FUNCTION_BLOCK FB 500
VERSION : 0.1


VAR_INPUT
  IN0 : BOOL ;
  IN1 : BOOL ;
  IN2 : BOOL ;
END_VAR
VAR_OUTPUT
  OUT3 : BOOL ;
  OUT4 : BOOL ;
END_VAR
VAR
  STAT5 : BOOL ;
  STAT6 : BOOL ;
  STAT7 : BOOL ;
  STAT8 : BOOL ;
END_VAR
BEGIN
NETWORK
TITLE =
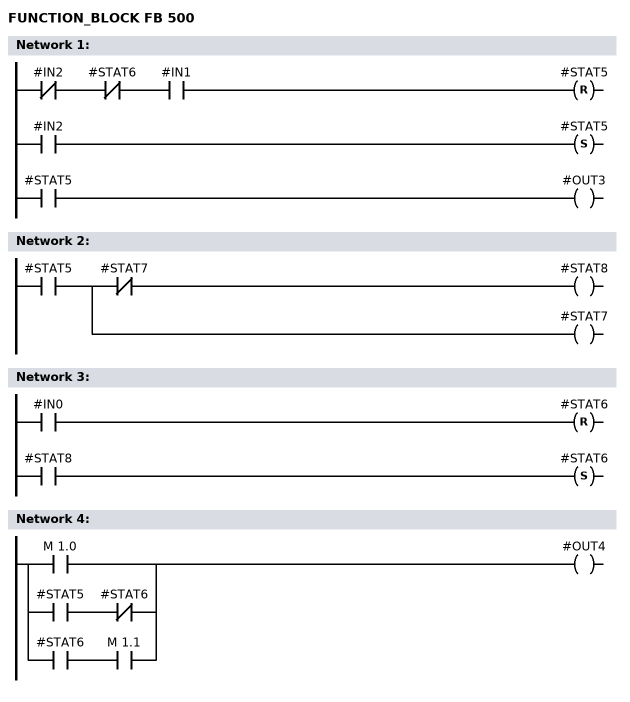

      AN    #IN2;
      AN    #STAT6;
      A     #IN1;
      R     #STAT5;
      A     #IN2;
      S     #STAT5;
      A     #STAT5;
      =     #OUT3;
NETWORK
TITLE =

      A     #STAT5;
      =     L      0.0;
      A     L      0.0;
      AN    #STAT7;
      =     #STAT8;
      A     L      0.0;
      BLD   102;
      =     #STAT7;
NETWORK
TITLE =

      A     #IN0;
      R     #STAT6;
      A     #STAT8;
      S     #STAT6;
      NOP   0;
NETWORK
TITLE =

      O     M      1.0;
      O     ;
      A     #STAT5;
      AN    #STAT6;
      O     ;
      A     #STAT6;
      A     M      1.1;
      =     #OUT4;
END_FUNCTION_BLOCK

FUNCTION FC 0 : VOID
VERSION : 0.1

BEGIN
NETWORK
TITLE =
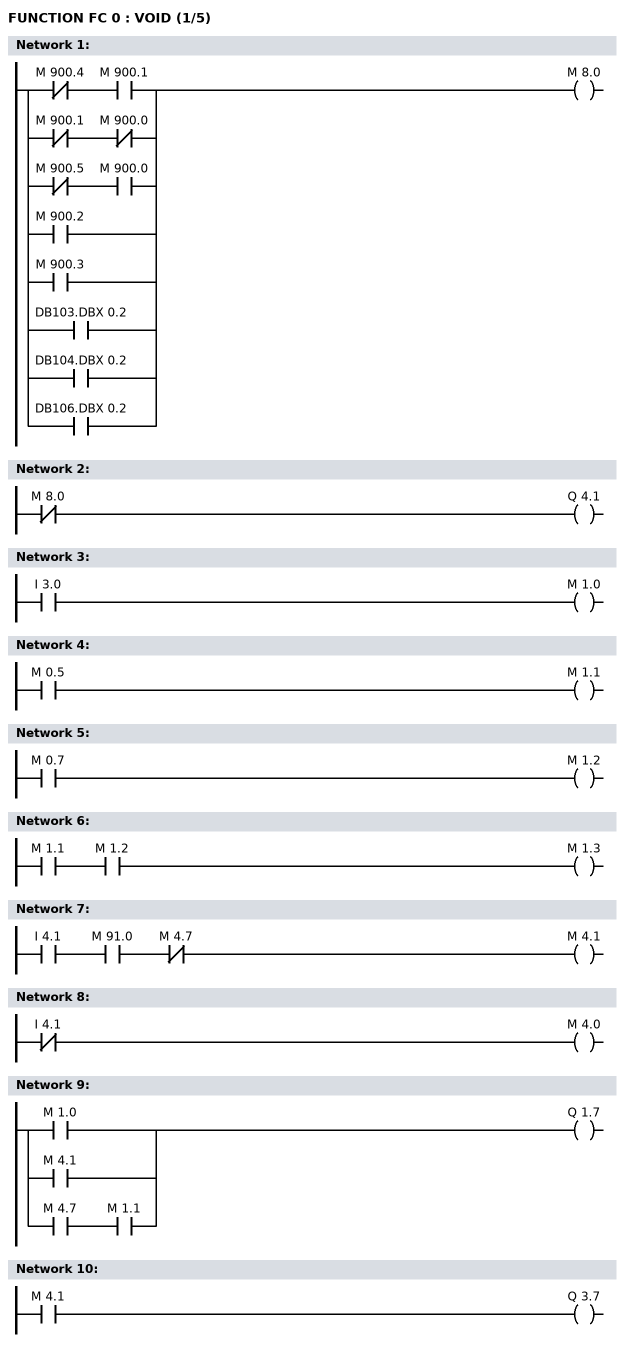

      AN    M    900.4;
      A     M    900.1;
      O     ;
      AN    M    900.1;
      AN    M    900.0;
      O     ;
      AN    M    900.5;
      A     M    900.0;
      O     M    900.2;
      O     M    900.3;
      O     DB103.DBX    0.2;
      O     DB104.DBX    0.2;
      O     DB106.DBX    0.2;
      =     M      8.0;
NETWORK
TITLE =

      AN    M      8.0;
      =     Q      4.1;
NETWORK
TITLE =

      A     I      3.0;
      =     M      1.0;
NETWORK
TITLE =

      A     M      0.5;
      =     M      1.1;
NETWORK
TITLE =

      A     M      0.7;
      =     M      1.2;
NETWORK
TITLE =

      A     M      1.1;
      A     M      1.2;
      =     M      1.3;
NETWORK
TITLE =

      A     I      4.1;
      A     M     91.0;
      AN    M      4.7;
      =     M      4.1;
NETWORK
TITLE =

      AN    I      4.1;
      =     M      4.0;
NETWORK
TITLE =

      O     M      1.0;
      O     M      4.1;
      O     ;
      A     M      4.7;
      A     M      1.1;
      =     Q      1.7;
NETWORK
TITLE =

      A     M      4.1;
      =     Q      3.7;
NETWORK
TITLE =
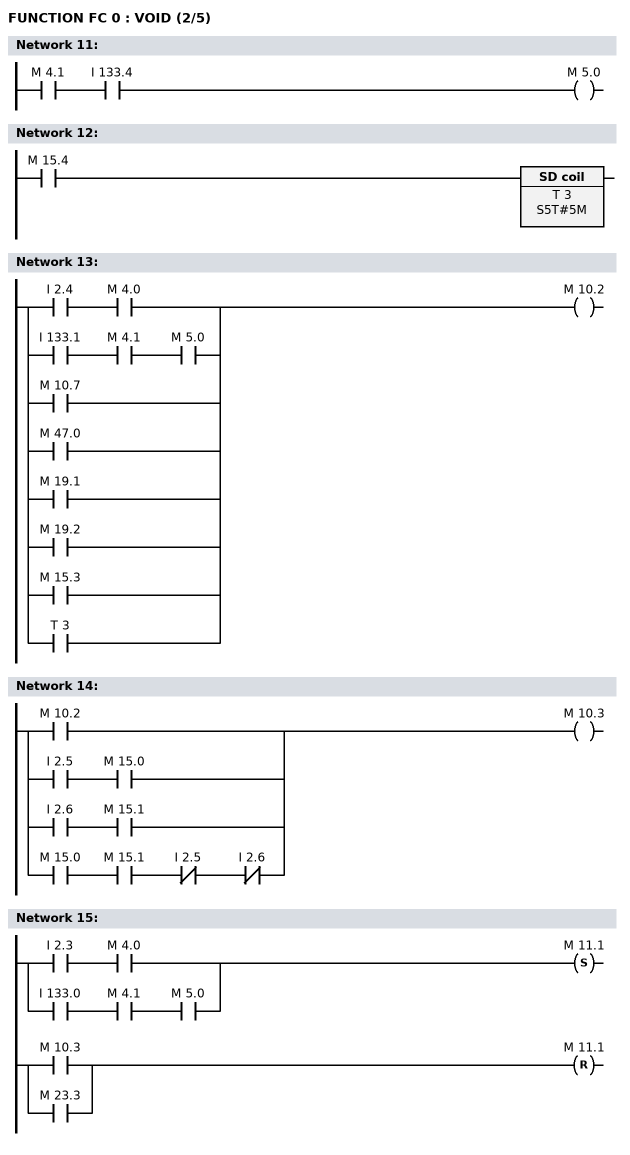

      A     M      4.1;
      A     I    133.4;
      =     M      5.0;
NETWORK
TITLE =

      A     M     15.4;
      L     S5T#5M;
      SD    T      3;
      NOP   0;
      NOP   0;
      NOP   0;
      NOP   0;
NETWORK
TITLE =

      A     I      2.4;
      A     M      4.0;
      O     ;
      A     I    133.1;
      A     M      4.1;
      A     M      5.0;
      O     M     10.7;
      O     M     47.0;
      O     M     19.1;
      O     M     19.2;
      O     M     15.3;
      O     T      3;
      =     M     10.2;
NETWORK
TITLE =

      O     M     10.2;
      O     ;
      A     I      2.5;
      A     M     15.0;
      O     ;
      A     I      2.6;
      A     M     15.1;
      O     ;
      A     M     15.0;
      A     M     15.1;
      AN    I      2.5;
      AN    I      2.6;
      =     M     10.3;
NETWORK
TITLE =

      A(    ;
      A     I      2.3;
      A     M      4.0;
      O     ;
      A     I    133.0;
      A     M      4.1;
      A     M      5.0;
      )     ;
      S     M     11.1;
      A(    ;
      O     M     10.3;
      O     M     23.3;
      )     ;
      R     M     11.1;
      NOP   0;
NETWORK
TITLE =
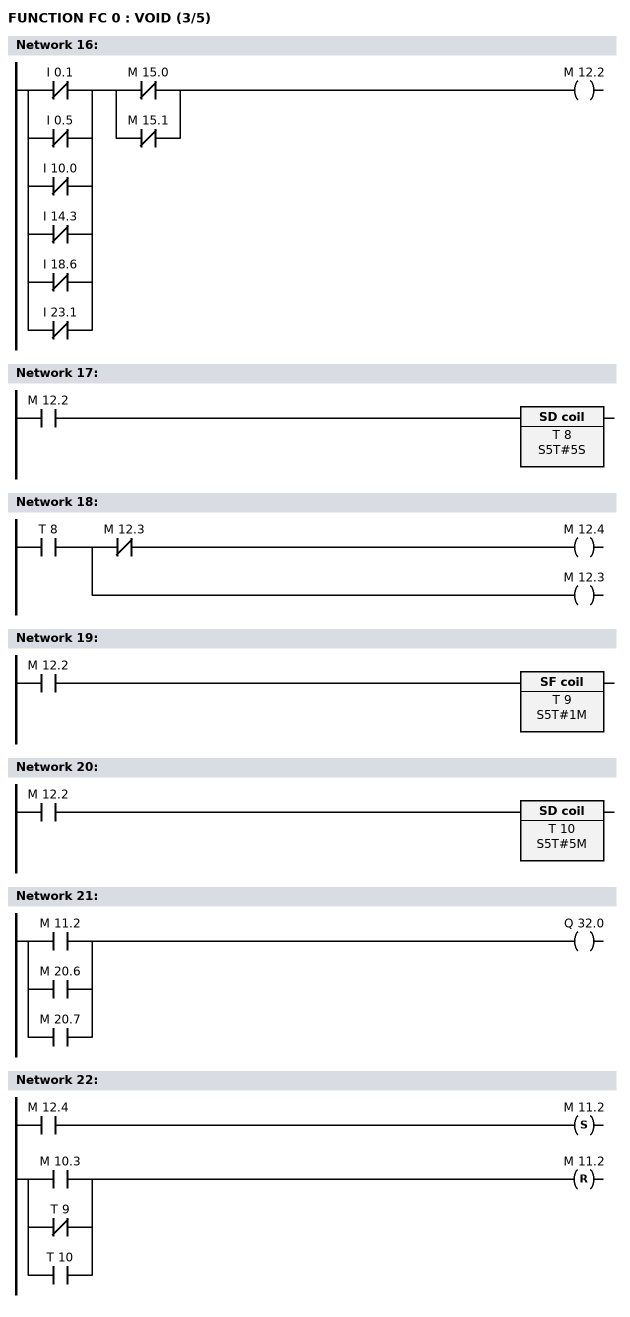

      A(    ;
      ON    I      0.1;
      ON    I      0.5;
      ON    I     10.0;
      ON    I     14.3;
      ON    I     18.6;
      ON    I     23.1;
      )     ;
      A(    ;
      ON    M     15.0;
      ON    M     15.1;
      )     ;
      =     M     12.2;
NETWORK
TITLE =

      A     M     12.2;
      L     S5T#5S;
      SD    T      8;
      NOP   0;
      NOP   0;
      NOP   0;
      NOP   0;
NETWORK
TITLE =

      A     T      8;
      =     L      0.0;
      A     L      0.0;
      AN    M     12.3;
      =     M     12.4;
      A     L      0.0;
      BLD   102;
      =     M     12.3;
NETWORK
TITLE =

      A     M     12.2;
      L     S5T#1M;
      SF    T      9;
      NOP   0;
      NOP   0;
      NOP   0;
      NOP   0;
NETWORK
TITLE =

      A     M     12.2;
      L     S5T#5M;
      SD    T     10;
      NOP   0;
      NOP   0;
      NOP   0;
      NOP   0;
NETWORK
TITLE =

      O     M     11.2;
      O     M     20.6;
      O     M     20.7;
      =     Q     32.0;
NETWORK
TITLE =

      A     M     12.4;
      S     M     11.2;
      A(    ;
      O     M     10.3;
      ON    T      9;
      O     T     10;
      )     ;
      R     M     11.2;
      NOP   0;
NETWORK
TITLE =
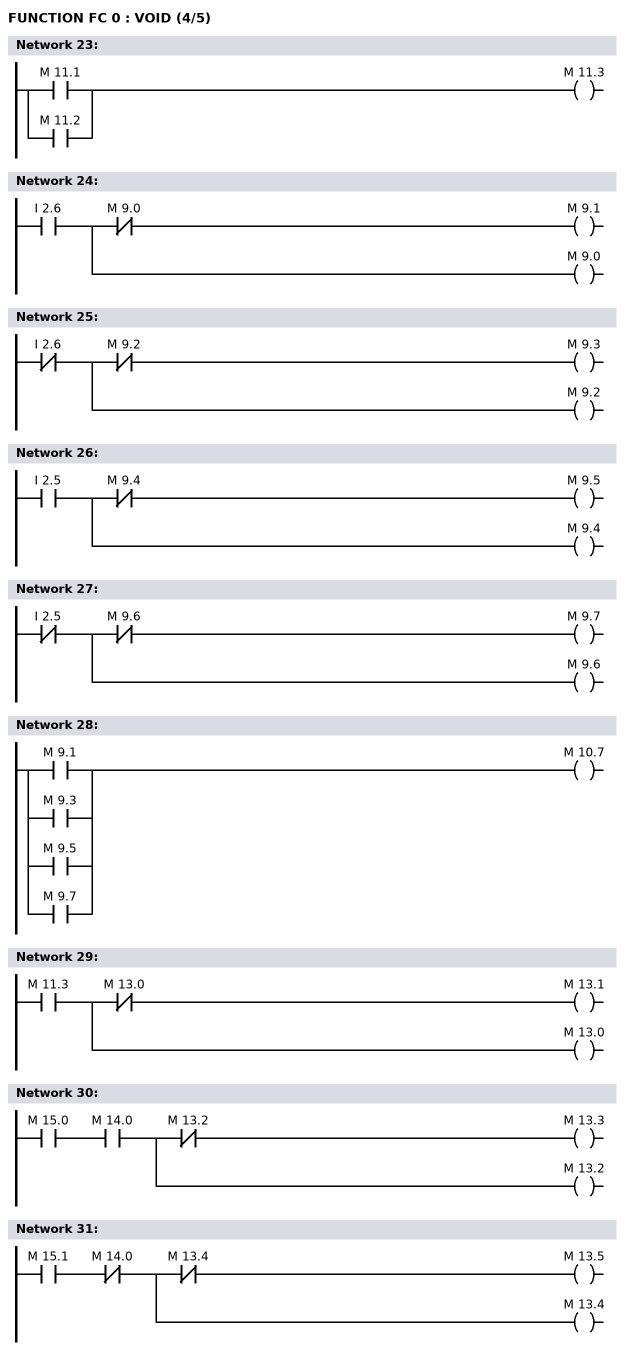

      O     M     11.1;
      O     M     11.2;
      =     M     11.3;
NETWORK
TITLE =

      A     I      2.6;
      =     L      0.0;
      A     L      0.0;
      AN    M      9.0;
      =     M      9.1;
      A     L      0.0;
      BLD   102;
      =     M      9.0;
NETWORK
TITLE =

      AN    I      2.6;
      =     L      0.0;
      A     L      0.0;
      AN    M      9.2;
      =     M      9.3;
      A     L      0.0;
      BLD   102;
      =     M      9.2;
NETWORK
TITLE =

      A     I      2.5;
      =     L      0.0;
      A     L      0.0;
      AN    M      9.4;
      =     M      9.5;
      A     L      0.0;
      BLD   102;
      =     M      9.4;
NETWORK
TITLE =

      AN    I      2.5;
      =     L      0.0;
      A     L      0.0;
      AN    M      9.6;
      =     M      9.7;
      A     L      0.0;
      BLD   102;
      =     M      9.6;
NETWORK
TITLE =

      O     M      9.1;
      O     M      9.3;
      O     M      9.5;
      O     M      9.7;
      =     M     10.7;
NETWORK
TITLE =

      A     M     11.3;
      =     L      0.0;
      A     L      0.0;
      AN    M     13.0;
      =     M     13.1;
      A     L      0.0;
      BLD   102;
      =     M     13.0;
NETWORK
TITLE =

      A     M     15.0;
      A     M     14.0;
      =     L      0.0;
      A     L      0.0;
      AN    M     13.2;
      =     M     13.3;
      A     L      0.0;
      BLD   102;
      =     M     13.2;
NETWORK
TITLE =

      A     M     15.1;
      AN    M     14.0;
      =     L      0.0;
      A     L      0.0;
      AN    M     13.4;
      =     M     13.5;
      A     L      0.0;
      BLD   102;
      =     M     13.4;
NETWORK
TITLE =
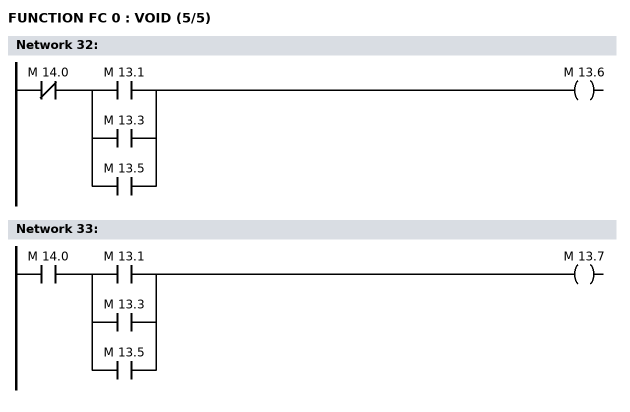

      AN    M     14.0;
      A(    ;
      O     M     13.1;
      O     M     13.3;
      O     M     13.5;
      )     ;
      =     M     13.6;
NETWORK
TITLE =

      A     M     14.0;
      A(    ;
      O     M     13.1;
      O     M     13.3;
      O     M     13.5;
      )     ;
      =     M     13.7;
NETWORK
TITLE =

      A(    ;
      A     M     13.7;
      R     M     14.0;
      A     M     13.6;
      S     M     14.0;
      A     M     14.0;
      )     ;
      AN    I      2.5;
      AN    I      2.6;
      O     I      2.5;
      =     M     14.2;
NETWORK
TITLE =
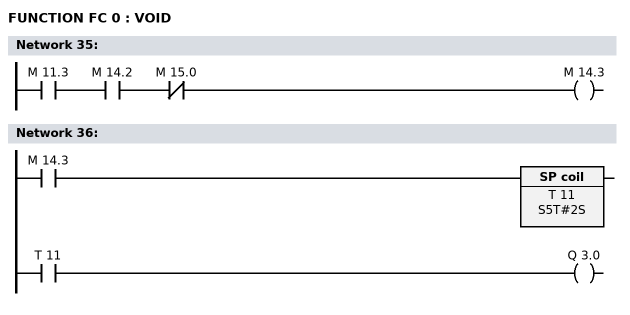

      A     M     11.3;
      A     M     14.2;
      AN    M     15.0;
      =     M     14.3;
NETWORK
TITLE =

      A     M     14.3;
      L     S5T#2S;
      SP    T     11;
      NOP   0;
      NOP   0;
      NOP   0;
      A     T     11;
      =     Q      3.0;
NETWORK
TITLE =

      A(    ;
      AN    M     14.3;
      L     S5T#2S;
      SP    T     12;
      NOP   0;
      NOP   0;
      NOP   0;
      A     T     12;
      )     ;
      NOT   ;
      =     Q      3.1;
NETWORK
TITLE =
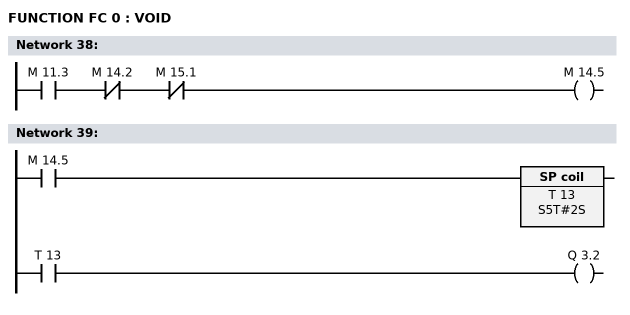

      A     M     11.3;
      AN    M     14.2;
      AN    M     15.1;
      =     M     14.5;
NETWORK
TITLE =

      A     M     14.5;
      L     S5T#2S;
      SP    T     13;
      NOP   0;
      NOP   0;
      NOP   0;
      A     T     13;
      =     Q      3.2;
NETWORK
TITLE =

      A(    ;
      AN    M     14.5;
      L     S5T#2S;
      SP    T     14;
      NOP   0;
      NOP   0;
      NOP   0;
      A     T     14;
      )     ;
      NOT   ;
      =     Q      3.3;
NETWORK
TITLE =
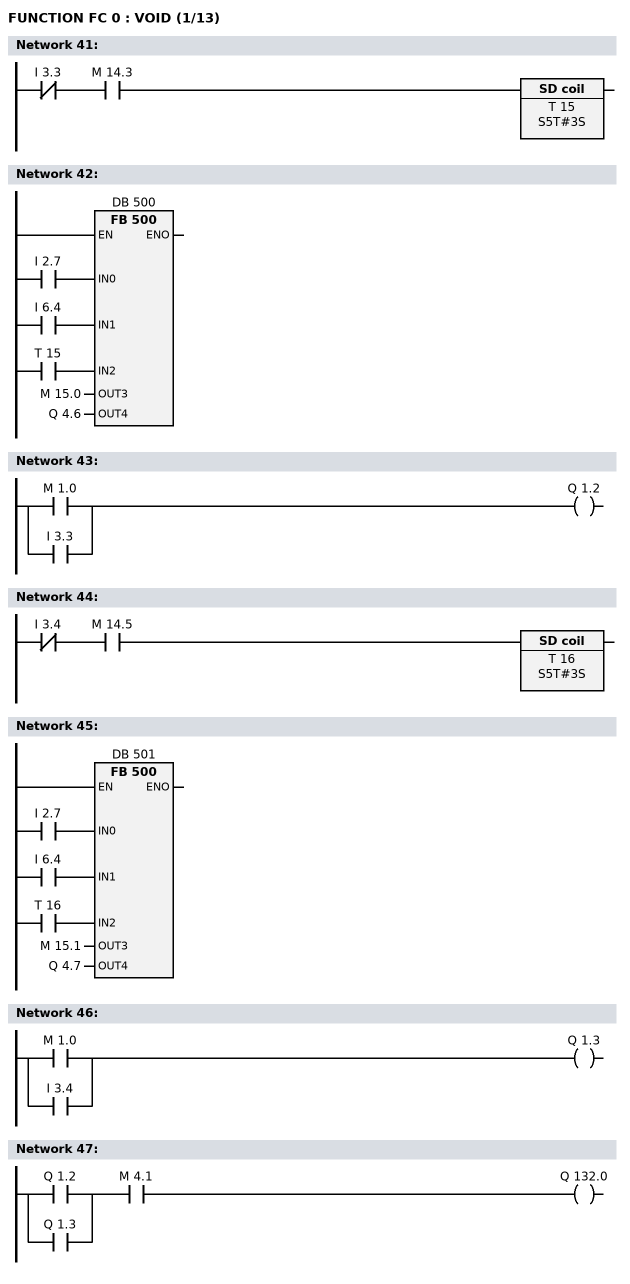

      AN    I      3.3;
      A     M     14.3;
      L     S5T#3S;
      SD    T     15;
      NOP   0;
      NOP   0;
      NOP   0;
      NOP   0;
NETWORK
TITLE =

      A     I      2.7;
      =     L      0.0;
      BLD   103;
      A     I      6.4;
      =     L      0.1;
      BLD   103;
      A     T     15;
      =     L      0.2;
      BLD   103;
      CALL FB   500 , DB   500 (
           IN0                      := L      0.0,
           IN1                      := L      0.1,
           IN2                      := L      0.2,
           OUT3                     := M     15.0,
           OUT4                     := Q      4.6);
      NOP   0;
NETWORK
TITLE =

      O     M      1.0;
      O     I      3.3;
      =     Q      1.2;
NETWORK
TITLE =

      AN    I      3.4;
      A     M     14.5;
      L     S5T#3S;
      SD    T     16;
      NOP   0;
      NOP   0;
      NOP   0;
      NOP   0;
NETWORK
TITLE =

      A     I      2.7;
      =     L      0.0;
      BLD   103;
      A     I      6.4;
      =     L      0.1;
      BLD   103;
      A     T     16;
      =     L      0.2;
      BLD   103;
      CALL FB   500 , DB   501 (
           IN0                      := L      0.0,
           IN1                      := L      0.1,
           IN2                      := L      0.2,
           OUT3                     := M     15.1,
           OUT4                     := Q      4.7);
      NOP   0;
NETWORK
TITLE =

      O     M      1.0;
      O     I      3.4;
      =     Q      1.3;
NETWORK
TITLE =

      A(    ;
      O     Q      1.2;
      O     Q      1.3;
      )     ;
      A     M      4.1;
      =     Q    132.0;
NETWORK
TITLE =
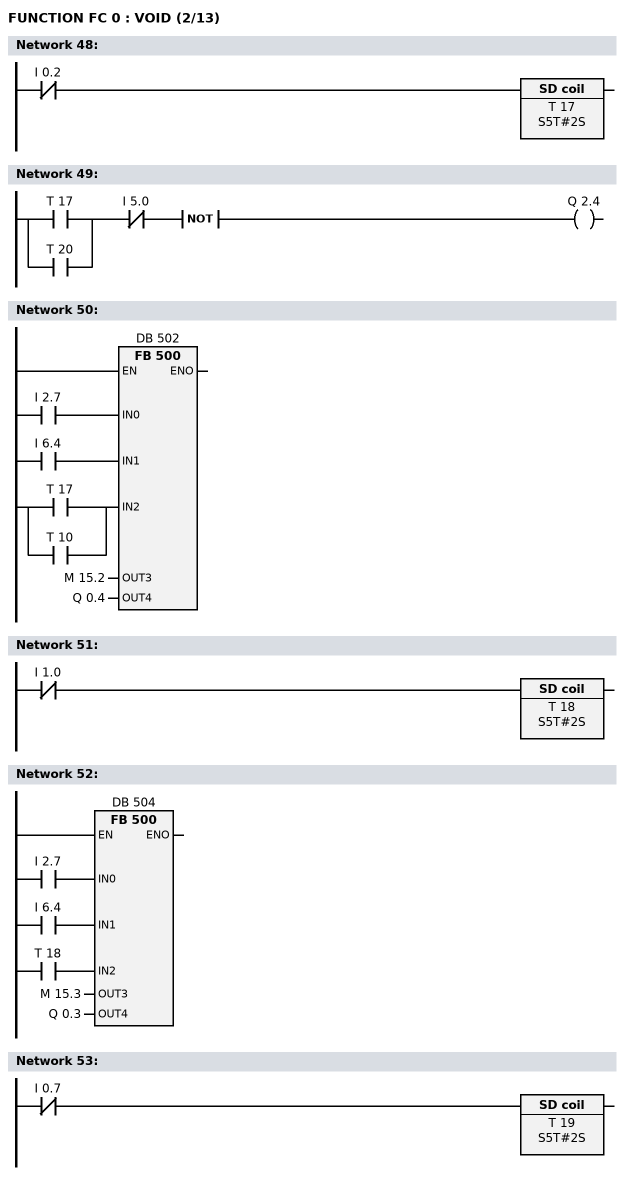

      AN    I      0.2;
      L     S5T#2S;
      SD    T     17;
      NOP   0;
      NOP   0;
      NOP   0;
      NOP   0;
NETWORK
TITLE =

      A(    ;
      O     T     17;
      O     T     20;
      )     ;
      AN    I      5.0;
      NOT   ;
      =     Q      2.4;
NETWORK
TITLE =

      A     I      2.7;
      =     L      0.0;
      BLD   103;
      A     I      6.4;
      =     L      0.1;
      BLD   103;
      A(    ;
      O     T     17;
      O     T     10;
      )     ;
      =     L      0.2;
      BLD   103;
      CALL FB   500 , DB   502 (
           IN0                      := L      0.0,
           IN1                      := L      0.1,
           IN2                      := L      0.2,
           OUT3                     := M     15.2,
           OUT4                     := Q      0.4);
      NOP   0;
NETWORK
TITLE =

      AN    I      1.0;
      L     S5T#2S;
      SD    T     18;
      NOP   0;
      NOP   0;
      NOP   0;
      NOP   0;
NETWORK
TITLE =

      A     I      2.7;
      =     L      0.0;
      BLD   103;
      A     I      6.4;
      =     L      0.1;
      BLD   103;
      A     T     18;
      =     L      0.2;
      BLD   103;
      CALL FB   500 , DB   504 (
           IN0                      := L      0.0,
           IN1                      := L      0.1,
           IN2                      := L      0.2,
           OUT3                     := M     15.3,
           OUT4                     := Q      0.3);
      NOP   0;
NETWORK
TITLE =

      AN    I      0.7;
      L     S5T#2S;
      SD    T     19;
      NOP   0;
      NOP   0;
      NOP   0;
      NOP   0;
NETWORK
TITLE =
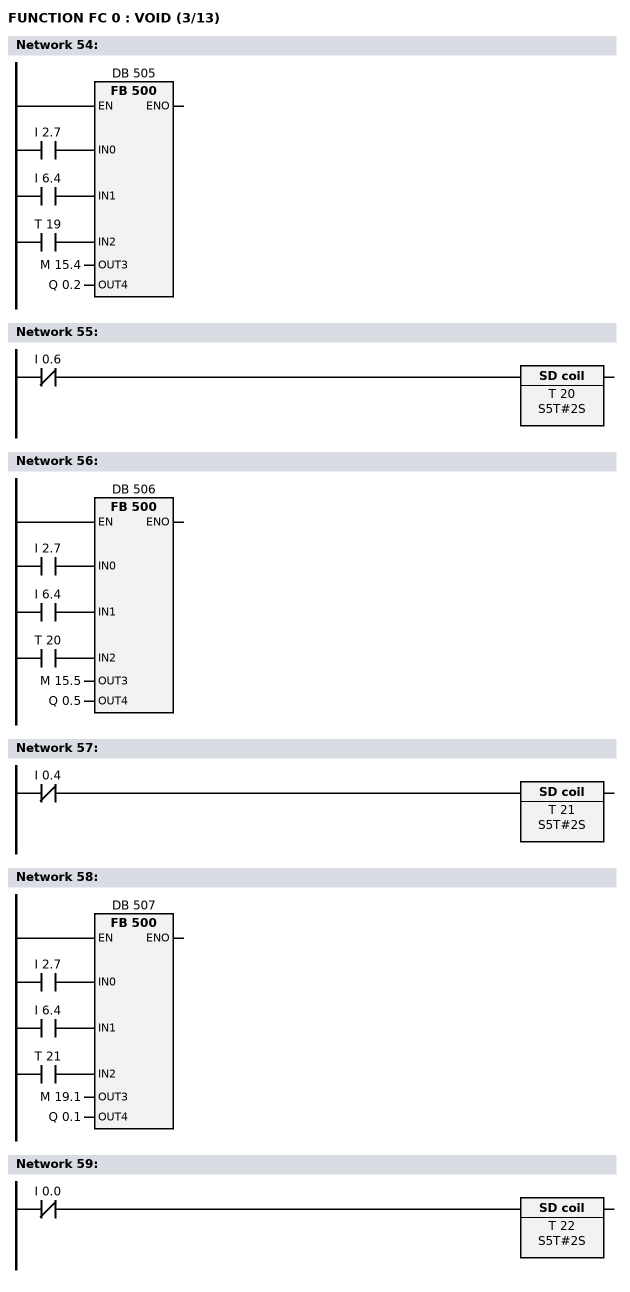

      A     I      2.7;
      =     L      0.0;
      BLD   103;
      A     I      6.4;
      =     L      0.1;
      BLD   103;
      A     T     19;
      =     L      0.2;
      BLD   103;
      CALL FB   500 , DB   505 (
           IN0                      := L      0.0,
           IN1                      := L      0.1,
           IN2                      := L      0.2,
           OUT3                     := M     15.4,
           OUT4                     := Q      0.2);
      NOP   0;
NETWORK
TITLE =

      AN    I      0.6;
      L     S5T#2S;
      SD    T     20;
      NOP   0;
      NOP   0;
      NOP   0;
      NOP   0;
NETWORK
TITLE =

      A     I      2.7;
      =     L      0.0;
      BLD   103;
      A     I      6.4;
      =     L      0.1;
      BLD   103;
      A     T     20;
      =     L      0.2;
      BLD   103;
      CALL FB   500 , DB   506 (
           IN0                      := L      0.0,
           IN1                      := L      0.1,
           IN2                      := L      0.2,
           OUT3                     := M     15.5,
           OUT4                     := Q      0.5);
      NOP   0;
NETWORK
TITLE =

      AN    I      0.4;
      L     S5T#2S;
      SD    T     21;
      NOP   0;
      NOP   0;
      NOP   0;
      NOP   0;
NETWORK
TITLE =

      A     I      2.7;
      =     L      0.0;
      BLD   103;
      A     I      6.4;
      =     L      0.1;
      BLD   103;
      A     T     21;
      =     L      0.2;
      BLD   103;
      CALL FB   500 , DB   507 (
           IN0                      := L      0.0,
           IN1                      := L      0.1,
           IN2                      := L      0.2,
           OUT3                     := M     19.1,
           OUT4                     := Q      0.1);
      NOP   0;
NETWORK
TITLE =

      AN    I      0.0;
      L     S5T#2S;
      SD    T     22;
      NOP   0;
      NOP   0;
      NOP   0;
      NOP   0;
NETWORK
TITLE =
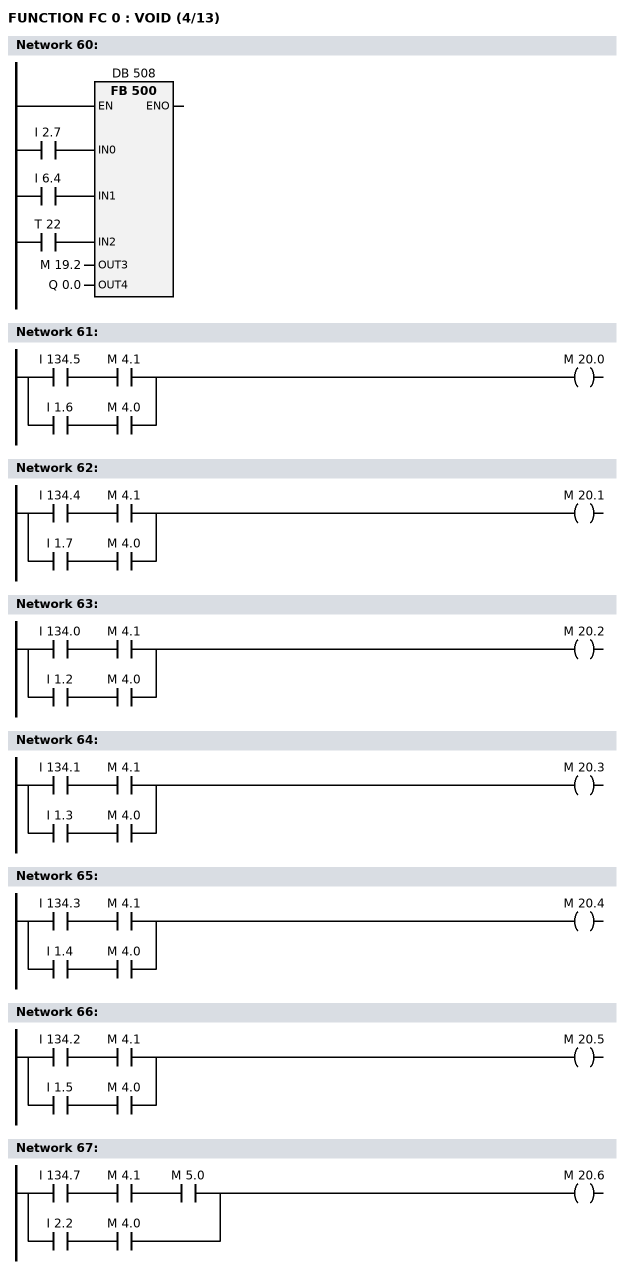

      A     I      2.7;
      =     L      0.0;
      BLD   103;
      A     I      6.4;
      =     L      0.1;
      BLD   103;
      A     T     22;
      =     L      0.2;
      BLD   103;
      CALL FB   500 , DB   508 (
           IN0                      := L      0.0,
           IN1                      := L      0.1,
           IN2                      := L      0.2,
           OUT3                     := M     19.2,
           OUT4                     := Q      0.0);
      NOP   0;
NETWORK
TITLE =

      A     I    134.5;
      A     M      4.1;
      O     ;
      A     I      1.6;
      A     M      4.0;
      =     M     20.0;
NETWORK
TITLE =

      A     I    134.4;
      A     M      4.1;
      O     ;
      A     I      1.7;
      A     M      4.0;
      =     M     20.1;
NETWORK
TITLE =

      A     I    134.0;
      A     M      4.1;
      O     ;
      A     I      1.2;
      A     M      4.0;
      =     M     20.2;
NETWORK
TITLE =

      A     I    134.1;
      A     M      4.1;
      O     ;
      A     I      1.3;
      A     M      4.0;
      =     M     20.3;
NETWORK
TITLE =

      A     I    134.3;
      A     M      4.1;
      O     ;
      A     I      1.4;
      A     M      4.0;
      =     M     20.4;
NETWORK
TITLE =

      A     I    134.2;
      A     M      4.1;
      O     ;
      A     I      1.5;
      A     M      4.0;
      =     M     20.5;
NETWORK
TITLE =

      A     I    134.7;
      A     M      4.1;
      A     M      5.0;
      O     ;
      A     I      2.2;
      A     M      4.0;
      =     M     20.6;
NETWORK
TITLE =
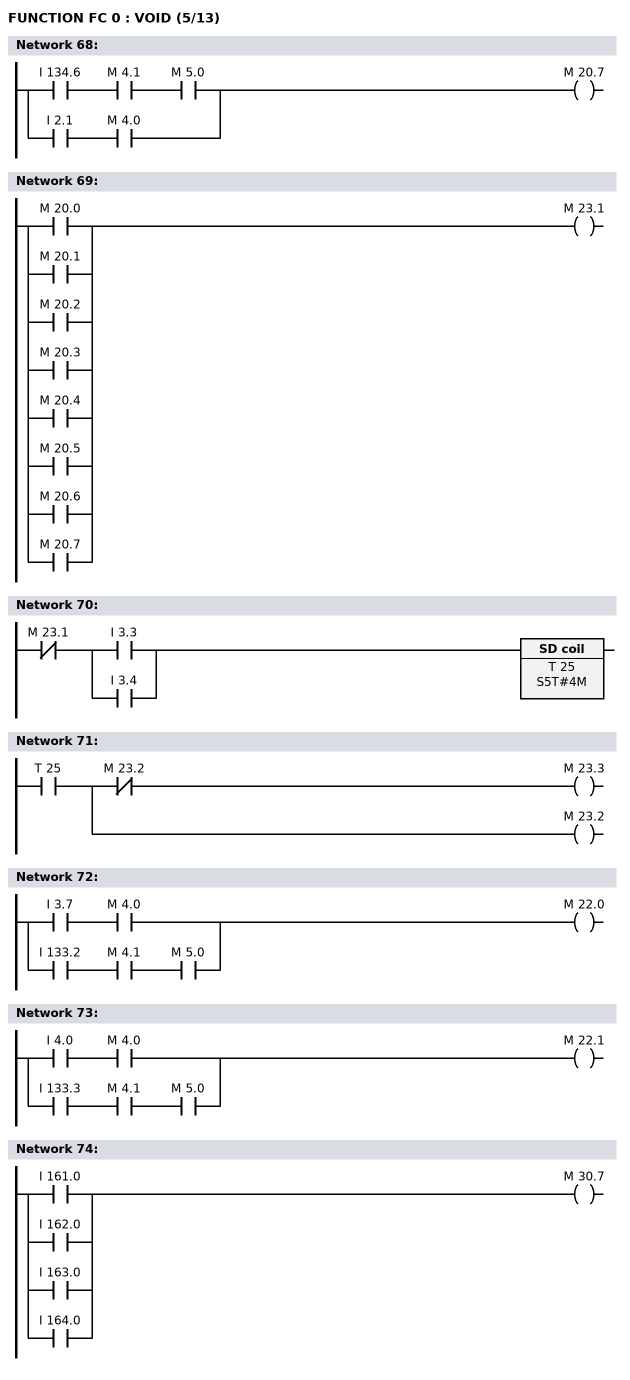

      A     I    134.6;
      A     M      4.1;
      A     M      5.0;
      O     ;
      A     I      2.1;
      A     M      4.0;
      =     M     20.7;
NETWORK
TITLE =

      O     M     20.0;
      O     M     20.1;
      O     M     20.2;
      O     M     20.3;
      O     M     20.4;
      O     M     20.5;
      O     M     20.6;
      O     M     20.7;
      =     M     23.1;
NETWORK
TITLE =

      AN    M     23.1;
      A(    ;
      O     I      3.3;
      O     I      3.4;
      )     ;
      L     S5T#4M;
      SD    T     25;
      NOP   0;
      NOP   0;
      NOP   0;
      NOP   0;
NETWORK
TITLE =

      A     T     25;
      =     L      0.0;
      A     L      0.0;
      AN    M     23.2;
      =     M     23.3;
      A     L      0.0;
      BLD   102;
      =     M     23.2;
NETWORK
TITLE =

      A     I      3.7;
      A     M      4.0;
      O     ;
      A     I    133.2;
      A     M      4.1;
      A     M      5.0;
      =     M     22.0;
NETWORK
TITLE =

      A     I      4.0;
      A     M      4.0;
      O     ;
      A     I    133.3;
      A     M      4.1;
      A     M      5.0;
      =     M     22.1;
NETWORK
TITLE =

      O     I    161.0;
      O     I    162.0;
      O     I    163.0;
      O     I    164.0;
      =     M     30.7;
NETWORK
TITLE =
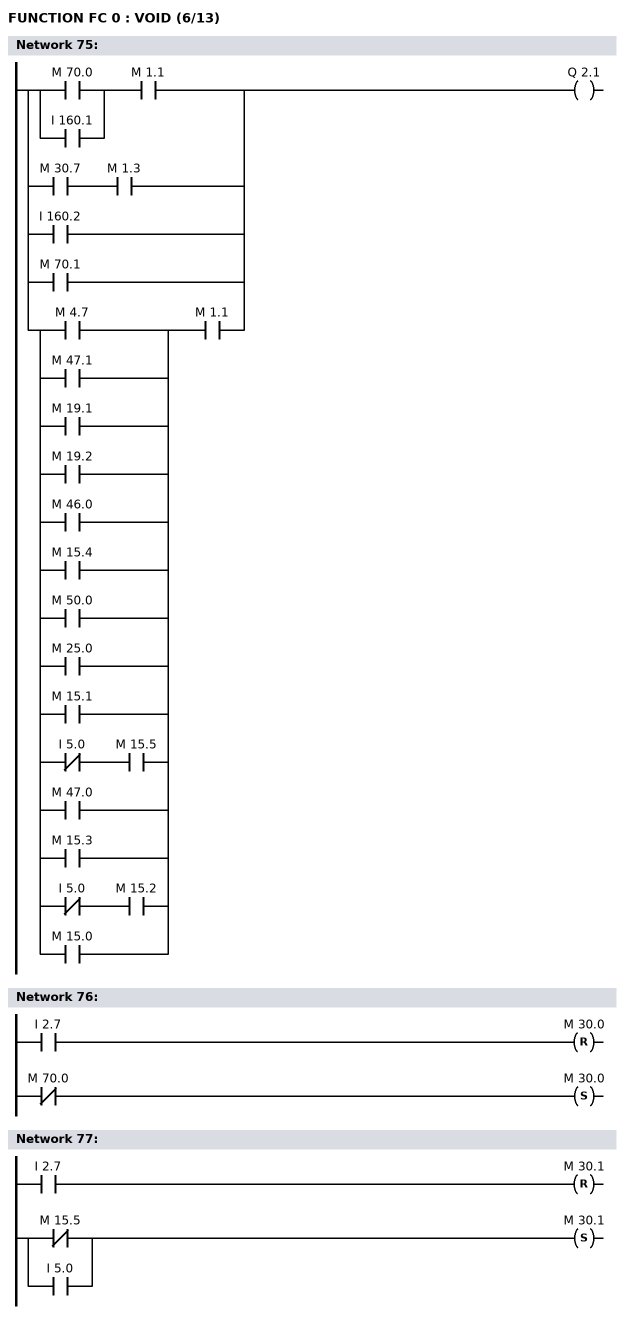

      A(    ;
      O     M     70.0;
      O     I    160.1;
      )     ;
      A     M      1.1;
      O     ;
      A     M     30.7;
      A     M      1.3;
      O     I    160.2;
      O     M     70.1;
      O     ;
      A(    ;
      O     M      4.7;
      O     M     47.1;
      O     M     19.1;
      O     M     19.2;
      O     M     46.0;
      O     M     15.4;
      O     M     50.0;
      O     M     25.0;
      O     M     15.1;
      O     ;
      AN    I      5.0;
      A     M     15.5;
      O     M     47.0;
      O     M     15.3;
      O     ;
      AN    I      5.0;
      A     M     15.2;
      O     M     15.0;
      )     ;
      A     M      1.1;
      =     Q      2.1;
NETWORK
TITLE =

      A     I      2.7;
      R     M     30.0;
      AN    M     70.0;
      S     M     30.0;
      NOP   0;
NETWORK
TITLE =

      A     I      2.7;
      R     M     30.1;
      A(    ;
      ON    M     15.5;
      O     I      5.0;
      )     ;
      S     M     30.1;
      NOP   0;
NETWORK
TITLE =
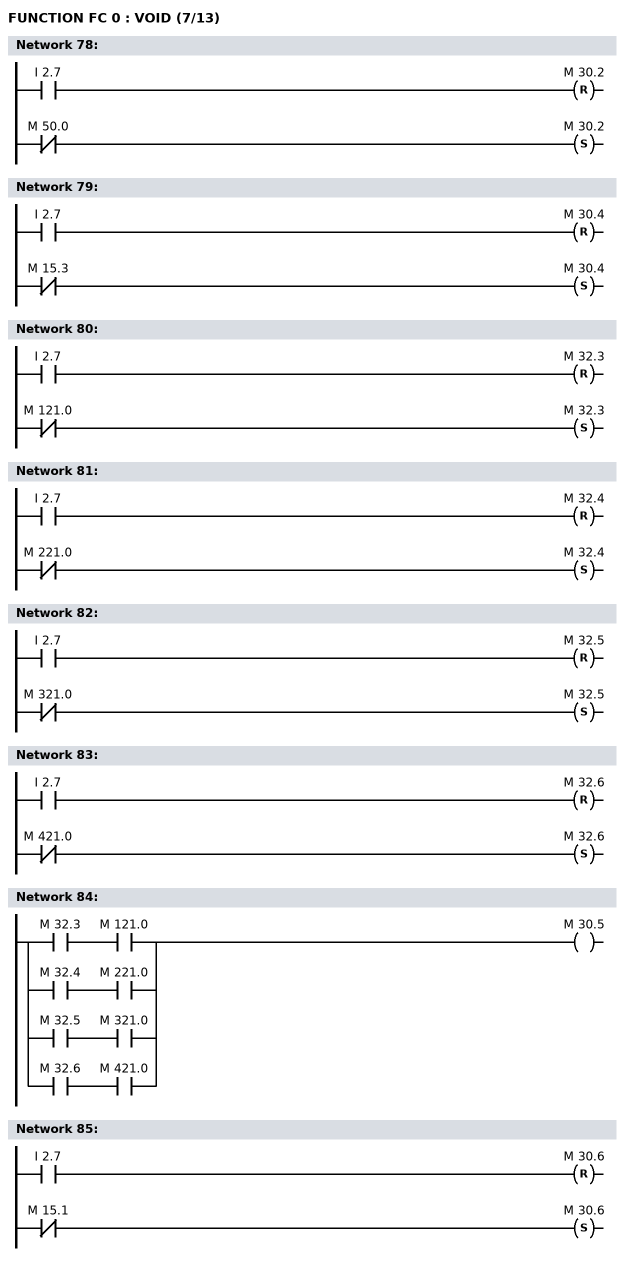

      A     I      2.7;
      R     M     30.2;
      AN    M     50.0;
      S     M     30.2;
      NOP   0;
NETWORK
TITLE =

      A     I      2.7;
      R     M     30.4;
      AN    M     15.3;
      S     M     30.4;
      NOP   0;
NETWORK
TITLE =

      A     I      2.7;
      R     M     32.3;
      AN    M    121.0;
      S     M     32.3;
      NOP   0;
NETWORK
TITLE =

      A     I      2.7;
      R     M     32.4;
      AN    M    221.0;
      S     M     32.4;
      NOP   0;
NETWORK
TITLE =

      A     I      2.7;
      R     M     32.5;
      AN    M    321.0;
      S     M     32.5;
      NOP   0;
NETWORK
TITLE =

      A     I      2.7;
      R     M     32.6;
      AN    M    421.0;
      S     M     32.6;
      NOP   0;
NETWORK
TITLE =

      A     M     32.3;
      A     M    121.0;
      O     ;
      A     M     32.4;
      A     M    221.0;
      O     ;
      A     M     32.5;
      A     M    321.0;
      O     ;
      A     M     32.6;
      A     M    421.0;
      =     M     30.5;
NETWORK
TITLE =

      A     I      2.7;
      R     M     30.6;
      AN    M     15.1;
      S     M     30.6;
      NOP   0;
NETWORK
TITLE =
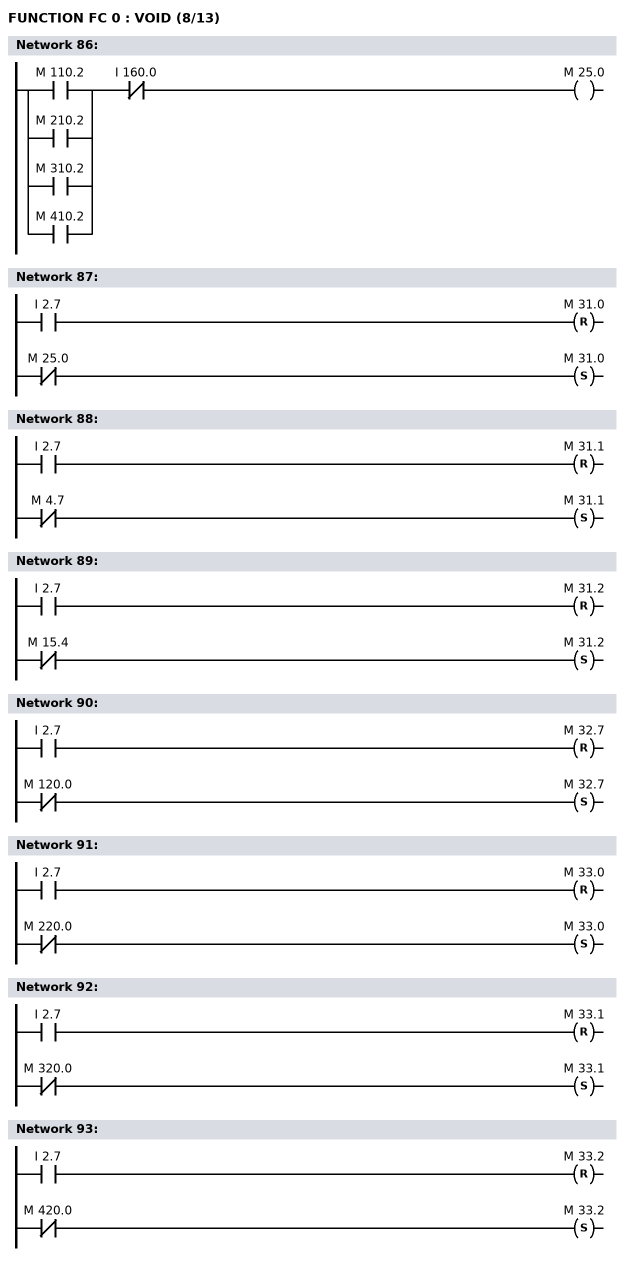

      A(    ;
      O     M    110.2;
      O     M    210.2;
      O     M    310.2;
      O     M    410.2;
      )     ;
      AN    I    160.0;
      =     M     25.0;
NETWORK
TITLE =

      A     I      2.7;
      R     M     31.0;
      AN    M     25.0;
      S     M     31.0;
      NOP   0;
NETWORK
TITLE =

      A     I      2.7;
      R     M     31.1;
      AN    M      4.7;
      S     M     31.1;
      NOP   0;
NETWORK
TITLE =

      A     I      2.7;
      R     M     31.2;
      AN    M     15.4;
      S     M     31.2;
      NOP   0;
NETWORK
TITLE =

      A     I      2.7;
      R     M     32.7;
      AN    M    120.0;
      S     M     32.7;
      NOP   0;
NETWORK
TITLE =

      A     I      2.7;
      R     M     33.0;
      AN    M    220.0;
      S     M     33.0;
      NOP   0;
NETWORK
TITLE =

      A     I      2.7;
      R     M     33.1;
      AN    M    320.0;
      S     M     33.1;
      NOP   0;
NETWORK
TITLE =

      A     I      2.7;
      R     M     33.2;
      AN    M    420.0;
      S     M     33.2;
      NOP   0;
NETWORK
TITLE =
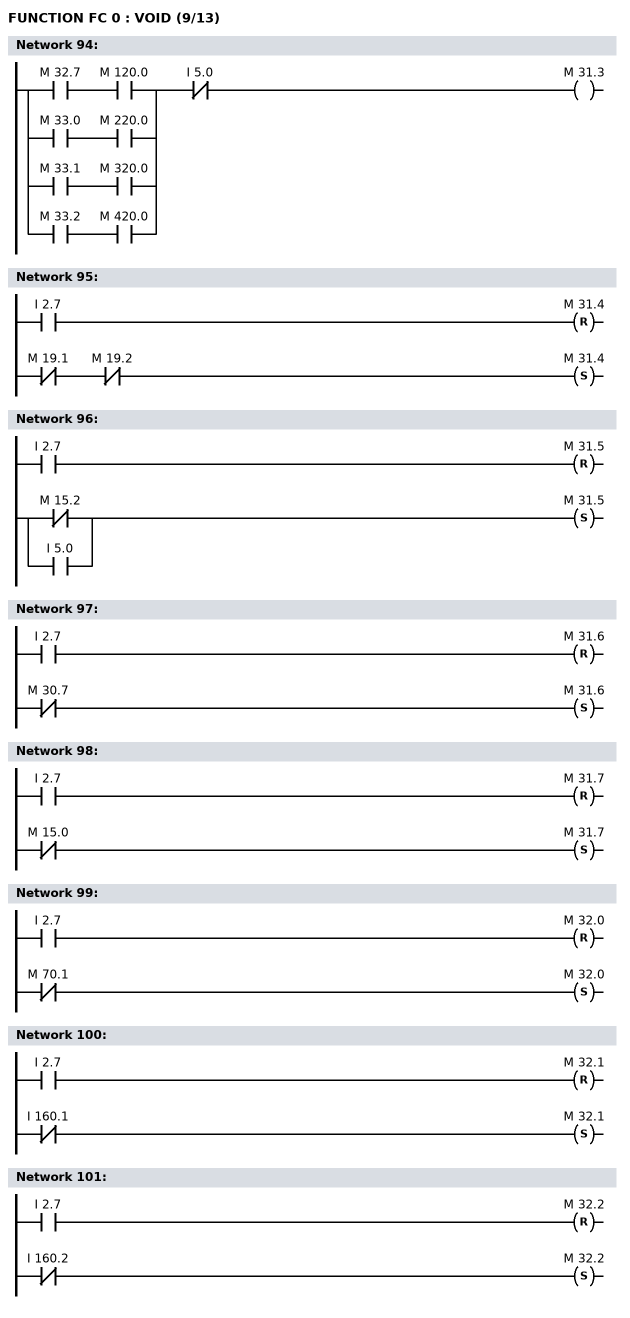

      A(    ;
      A     M     32.7;
      A     M    120.0;
      O     ;
      A     M     33.0;
      A     M    220.0;
      O     ;
      A     M     33.1;
      A     M    320.0;
      O     ;
      A     M     33.2;
      A     M    420.0;
      )     ;
      AN    I      5.0;
      =     M     31.3;
NETWORK
TITLE =

      A     I      2.7;
      R     M     31.4;
      AN    M     19.1;
      AN    M     19.2;
      S     M     31.4;
      NOP   0;
NETWORK
TITLE =

      A     I      2.7;
      R     M     31.5;
      A(    ;
      ON    M     15.2;
      O     I      5.0;
      )     ;
      S     M     31.5;
      NOP   0;
NETWORK
TITLE =

      A     I      2.7;
      R     M     31.6;
      AN    M     30.7;
      S     M     31.6;
      NOP   0;
NETWORK
TITLE =

      A     I      2.7;
      R     M     31.7;
      AN    M     15.0;
      S     M     31.7;
      NOP   0;
NETWORK
TITLE =

      A     I      2.7;
      R     M     32.0;
      AN    M     70.1;
      S     M     32.0;
      NOP   0;
NETWORK
TITLE =

      A     I      2.7;
      R     M     32.1;
      AN    I    160.1;
      S     M     32.1;
      NOP   0;
NETWORK
TITLE =

      A     I      2.7;
      R     M     32.2;
      AN    I    160.2;
      S     M     32.2;
      NOP   0;
NETWORK
TITLE =
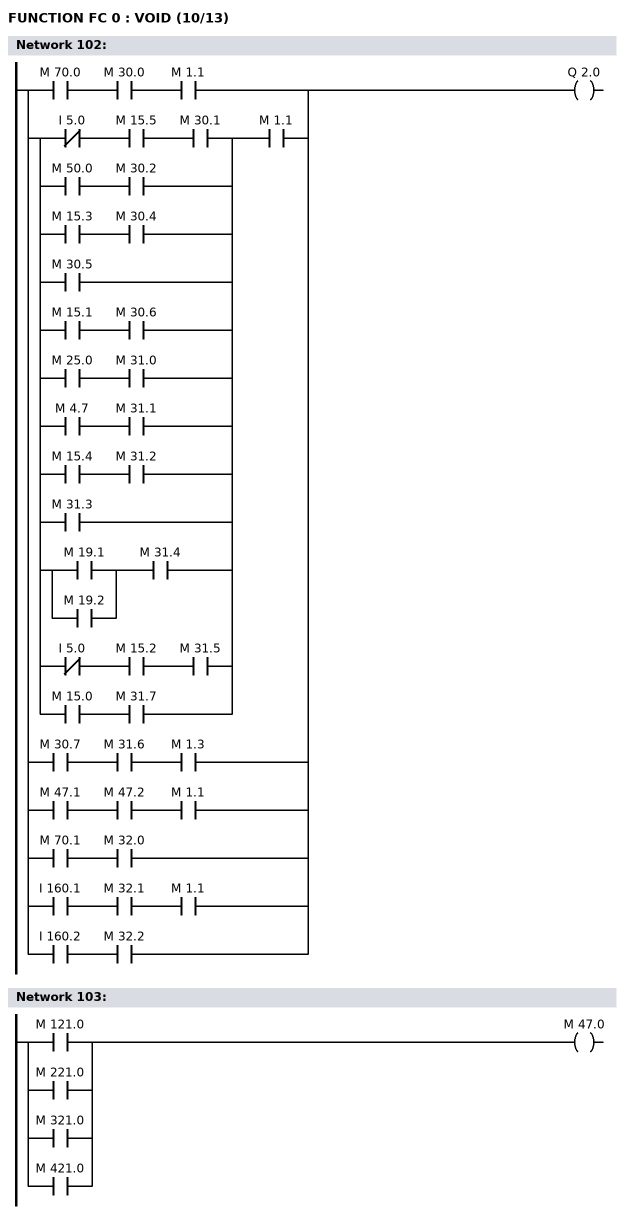

      A     M     70.0;
      A     M     30.0;
      A     M      1.1;
      O     ;
      A(    ;
      AN    I      5.0;
      A     M     15.5;
      A     M     30.1;
      O     ;
      A     M     50.0;
      A     M     30.2;
      O     ;
      A     M     15.3;
      A     M     30.4;
      O     M     30.5;
      O     ;
      A     M     15.1;
      A     M     30.6;
      O     ;
      A     M     25.0;
      A     M     31.0;
      O     ;
      A     M      4.7;
      A     M     31.1;
      O     ;
      A     M     15.4;
      A     M     31.2;
      O     M     31.3;
      O     ;
      A(    ;
      O     M     19.1;
      O     M     19.2;
      )     ;
      A     M     31.4;
      O     ;
      AN    I      5.0;
      A     M     15.2;
      A     M     31.5;
      O     ;
      A     M     15.0;
      A     M     31.7;
      )     ;
      A     M      1.1;
      O     ;
      A     M     30.7;
      A     M     31.6;
      A     M      1.3;
      O     ;
      A     M     47.1;
      A     M     47.2;
      A     M      1.1;
      O     ;
      A     M     70.1;
      A     M     32.0;
      O     ;
      A     I    160.1;
      A     M     32.1;
      A     M      1.1;
      O     ;
      A     I    160.2;
      A     M     32.2;
      =     Q      2.0;
NETWORK
TITLE =

      O     M    121.0;
      O     M    221.0;
      O     M    321.0;
      O     M    421.0;
      =     M     47.0;
NETWORK
TITLE =
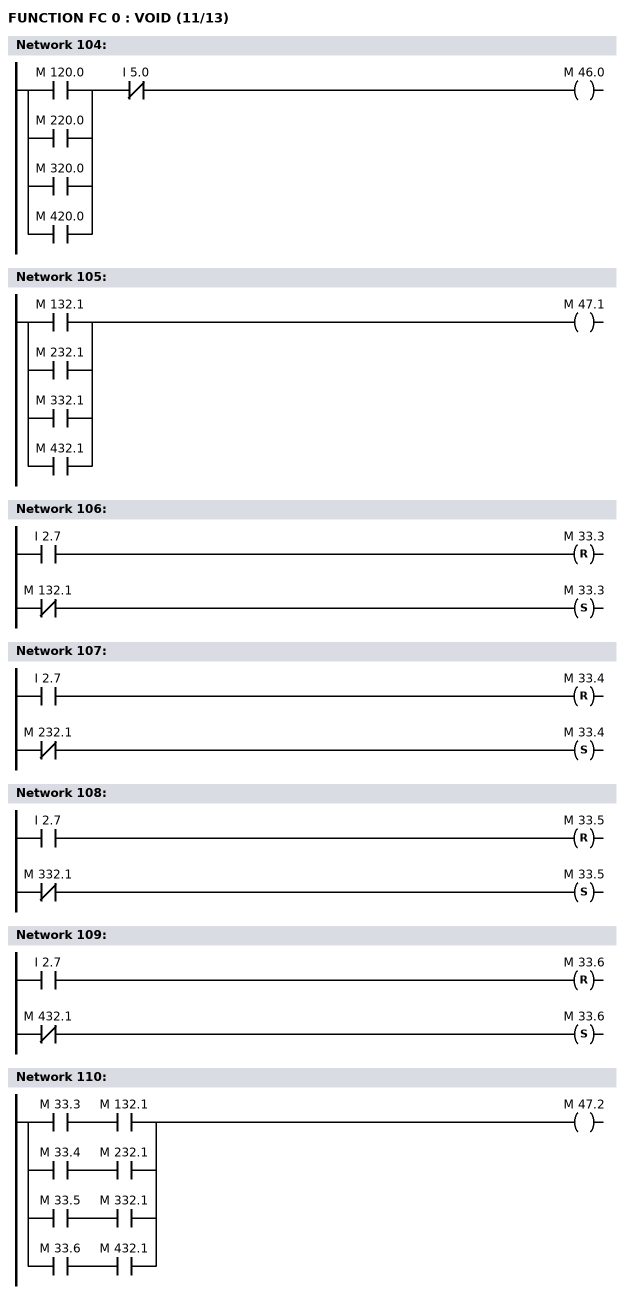

      A(    ;
      O     M    120.0;
      O     M    220.0;
      O     M    320.0;
      O     M    420.0;
      )     ;
      AN    I      5.0;
      =     M     46.0;
NETWORK
TITLE =

      O     M    132.1;
      O     M    232.1;
      O     M    332.1;
      O     M    432.1;
      =     M     47.1;
NETWORK
TITLE =

      A     I      2.7;
      R     M     33.3;
      AN    M    132.1;
      S     M     33.3;
      NOP   0;
NETWORK
TITLE =

      A     I      2.7;
      R     M     33.4;
      AN    M    232.1;
      S     M     33.4;
      NOP   0;
NETWORK
TITLE =

      A     I      2.7;
      R     M     33.5;
      AN    M    332.1;
      S     M     33.5;
      NOP   0;
NETWORK
TITLE =

      A     I      2.7;
      R     M     33.6;
      AN    M    432.1;
      S     M     33.6;
      NOP   0;
NETWORK
TITLE =

      A     M     33.3;
      A     M    132.1;
      O     ;
      A     M     33.4;
      A     M    232.1;
      O     ;
      A     M     33.5;
      A     M    332.1;
      O     ;
      A     M     33.6;
      A     M    432.1;
      =     M     47.2;
NETWORK
TITLE =
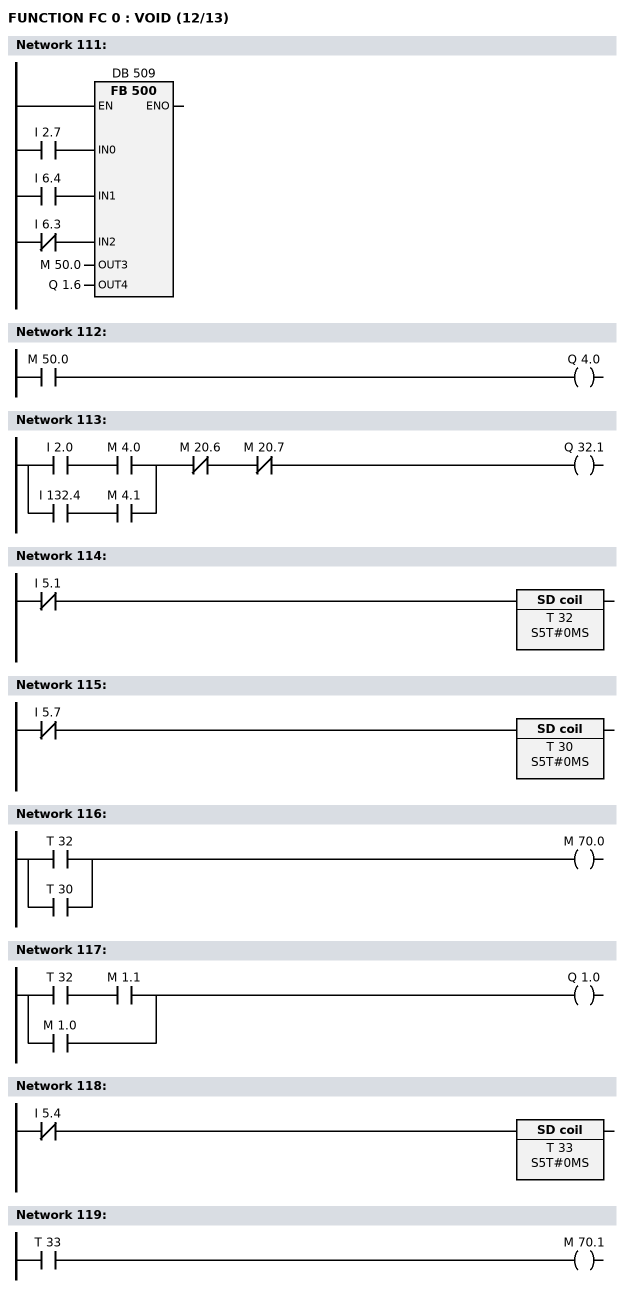

      A     I      2.7;
      =     L      0.0;
      BLD   103;
      A     I      6.4;
      =     L      0.1;
      BLD   103;
      AN    I      6.3;
      =     L      0.2;
      BLD   103;
      CALL FB   500 , DB   509 (
           IN0                      := L      0.0,
           IN1                      := L      0.1,
           IN2                      := L      0.2,
           OUT3                     := M     50.0,
           OUT4                     := Q      1.6);
      NOP   0;
NETWORK
TITLE =

      A     M     50.0;
      =     Q      4.0;
NETWORK
TITLE =

      A(    ;
      A     I      2.0;
      A     M      4.0;
      O     ;
      A     I    132.4;
      A     M      4.1;
      )     ;
      AN    M     20.6;
      AN    M     20.7;
      =     Q     32.1;
NETWORK
TITLE =

      AN    I      5.1;
      L     S5T#0MS;
      SD    T     32;
      NOP   0;
      NOP   0;
      NOP   0;
      NOP   0;
NETWORK
TITLE =

      AN    I      5.7;
      L     S5T#0MS;
      SD    T     30;
      NOP   0;
      NOP   0;
      NOP   0;
      NOP   0;
NETWORK
TITLE =

      O     T     32;
      O     T     30;
      =     M     70.0;
NETWORK
TITLE =

      A     T     32;
      A     M      1.1;
      O     M      1.0;
      =     Q      1.0;
NETWORK
TITLE =

      AN    I      5.4;
      L     S5T#0MS;
      SD    T     33;
      NOP   0;
      NOP   0;
      NOP   0;
      NOP   0;
NETWORK
TITLE =

      A     T     33;
      =     M     70.1;
NETWORK
TITLE =
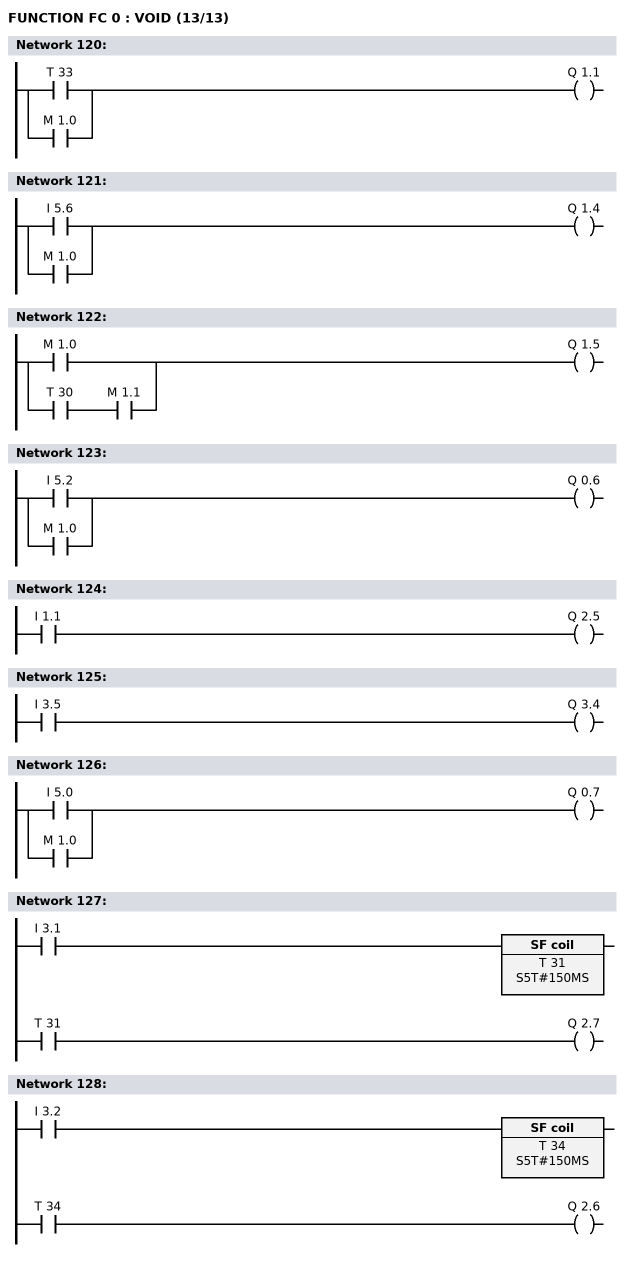

      O     T     33;
      O     M      1.0;
      =     Q      1.1;
NETWORK
TITLE =

      O     I      5.6;
      O     M      1.0;
      =     Q      1.4;
NETWORK
TITLE =

      O     M      1.0;
      O     ;
      A     T     30;
      A     M      1.1;
      =     Q      1.5;
NETWORK
TITLE =

      O     I      5.2;
      O     M      1.0;
      =     Q      0.6;
NETWORK
TITLE =

      A     I      1.1;
      =     Q      2.5;
NETWORK
TITLE =

      A     I      3.5;
      =     Q      3.4;
NETWORK
TITLE =

      O     I      5.0;
      O     M      1.0;
      =     Q      0.7;
NETWORK
TITLE =

      A     I      3.1;
      L     S5T#150MS;
      SF    T     31;
      NOP   0;
      NOP   0;
      NOP   0;
      A     T     31;
      =     Q      2.7;
NETWORK
TITLE =

      A     I      3.2;
      L     S5T#150MS;
      SF    T     34;
      NOP   0;
      NOP   0;
      NOP   0;
      A     T     34;
      =     Q      2.6;
END_FUNCTION

FUNCTION FC 1 : VOID
VERSION : 0.1

BEGIN
NETWORK
TITLE =
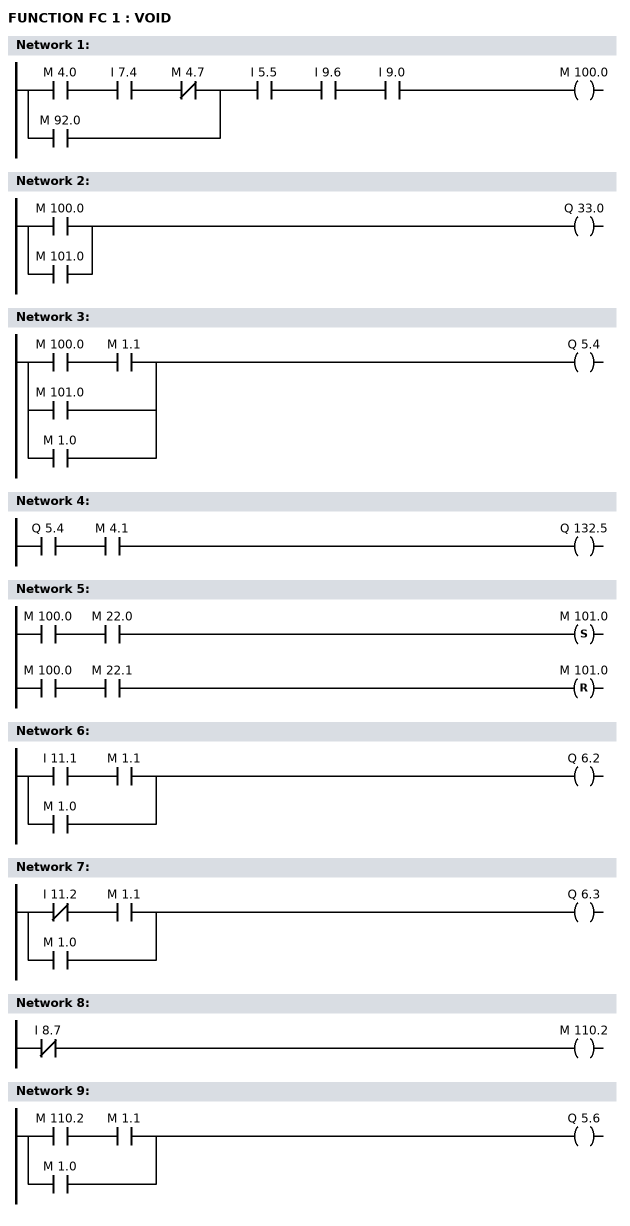

      A(    ;
      A     M      4.0;
      A     I      7.4;
      AN    M      4.7;
      O     M     92.0;
      )     ;
      A     I      5.5;
      A     I      9.6;
      A     I      9.0;
      =     M    100.0;
NETWORK
TITLE =

      O     M    100.0;
      O     M    101.0;
      =     Q     33.0;
NETWORK
TITLE =

      A     M    100.0;
      A     M      1.1;
      O     M    101.0;
      O     M      1.0;
      =     Q      5.4;
NETWORK
TITLE =

      A     Q      5.4;
      A     M      4.1;
      =     Q    132.5;
NETWORK
TITLE =

      A     M    100.0;
      A     M     22.0;
      S     M    101.0;
      A     M    100.0;
      A     M     22.1;
      R     M    101.0;
      NOP   0;
NETWORK
TITLE =

      A     I     11.1;
      A     M      1.1;
      O     M      1.0;
      =     Q      6.2;
NETWORK
TITLE =

      AN    I     11.2;
      A     M      1.1;
      O     M      1.0;
      =     Q      6.3;
NETWORK
TITLE =

      AN    I      8.7;
      =     M    110.2;
NETWORK
TITLE =

      A     M    110.2;
      A     M      1.1;
      O     M      1.0;
      =     Q      5.6;
NETWORK
TITLE =

      O(    ;
      A     I      8.0;
      L     S5T#150MS;
      SD    T     50;
      NOP   0;
      NOP   0;
      NOP   0;
      A     T     50;
      )     ;
      O     M      1.0;
      =     Q      5.3;
NETWORK
TITLE =
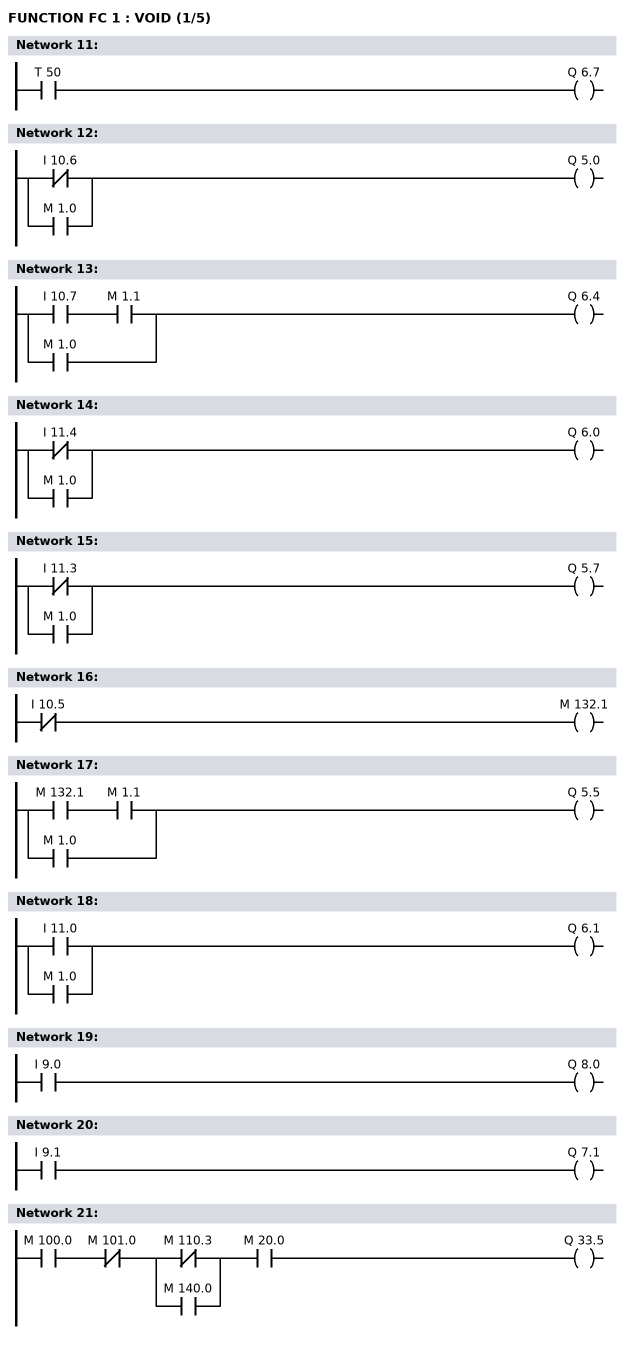

      A     T     50;
      =     Q      6.7;
NETWORK
TITLE =

      ON    I     10.6;
      O     M      1.0;
      =     Q      5.0;
NETWORK
TITLE =

      A     I     10.7;
      A     M      1.1;
      O     M      1.0;
      =     Q      6.4;
NETWORK
TITLE =

      ON    I     11.4;
      O     M      1.0;
      =     Q      6.0;
NETWORK
TITLE =

      ON    I     11.3;
      O     M      1.0;
      =     Q      5.7;
NETWORK
TITLE =

      AN    I     10.5;
      =     M    132.1;
NETWORK
TITLE =

      A     M    132.1;
      A     M      1.1;
      O     M      1.0;
      =     Q      5.5;
NETWORK
TITLE =

      O     I     11.0;
      O     M      1.0;
      =     Q      6.1;
NETWORK
TITLE =

      A     I      9.0;
      =     Q      8.0;
NETWORK
TITLE =

      A     I      9.1;
      =     Q      7.1;
NETWORK
TITLE =

      A     M    100.0;
      AN    M    101.0;
      A(    ;
      ON    M    110.3;
      O     M    140.0;
      )     ;
      A     M     20.0;
      =     Q     33.5;
NETWORK
TITLE =
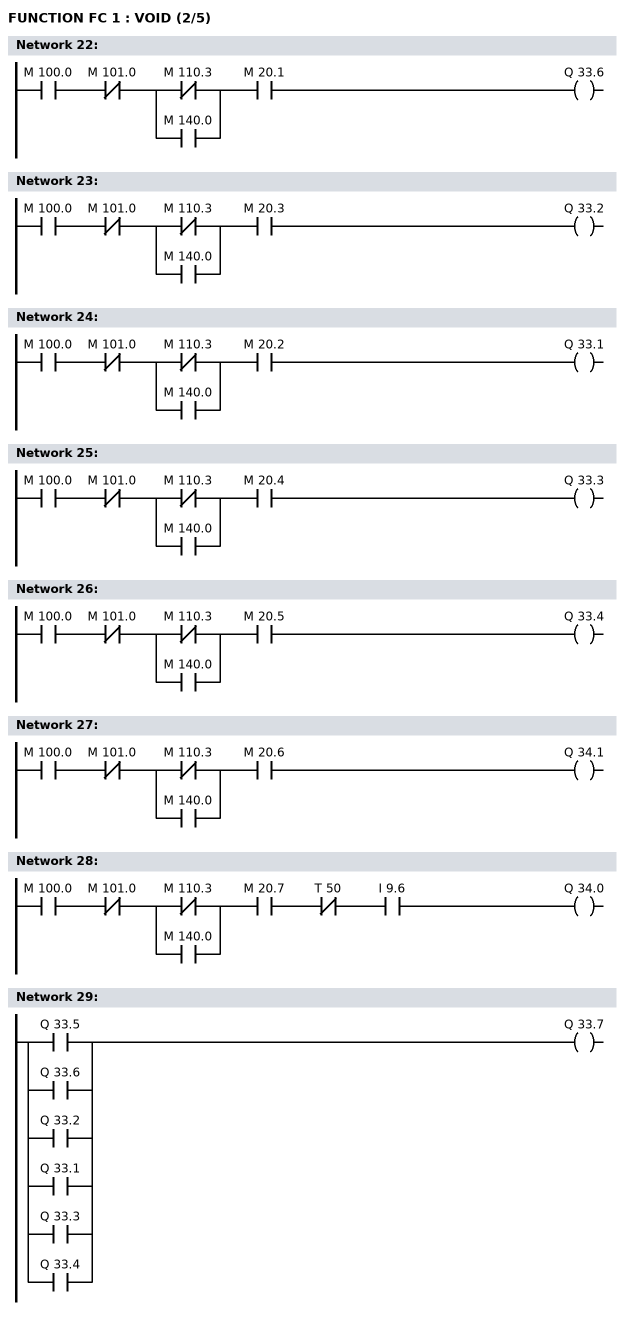

      A     M    100.0;
      AN    M    101.0;
      A(    ;
      ON    M    110.3;
      O     M    140.0;
      )     ;
      A     M     20.1;
      =     Q     33.6;
NETWORK
TITLE =

      A     M    100.0;
      AN    M    101.0;
      A(    ;
      ON    M    110.3;
      O     M    140.0;
      )     ;
      A     M     20.3;
      =     Q     33.2;
NETWORK
TITLE =

      A     M    100.0;
      AN    M    101.0;
      A(    ;
      ON    M    110.3;
      O     M    140.0;
      )     ;
      A     M     20.2;
      =     Q     33.1;
NETWORK
TITLE =

      A     M    100.0;
      AN    M    101.0;
      A(    ;
      ON    M    110.3;
      O     M    140.0;
      )     ;
      A     M     20.4;
      =     Q     33.3;
NETWORK
TITLE =

      A     M    100.0;
      AN    M    101.0;
      A(    ;
      ON    M    110.3;
      O     M    140.0;
      )     ;
      A     M     20.5;
      =     Q     33.4;
NETWORK
TITLE =

      A     M    100.0;
      AN    M    101.0;
      A(    ;
      ON    M    110.3;
      O     M    140.0;
      )     ;
      A     M     20.6;
      =     Q     34.1;
NETWORK
TITLE =

      A     M    100.0;
      AN    M    101.0;
      A(    ;
      ON    M    110.3;
      O     M    140.0;
      )     ;
      A     M     20.7;
      AN    T     50;
      A     I      9.6;
      =     Q     34.0;
NETWORK
TITLE =

      O     Q     33.5;
      O     Q     33.6;
      O     Q     33.2;
      O     Q     33.1;
      O     Q     33.3;
      O     Q     33.4;
      =     Q     33.7;
NETWORK
TITLE =
